Staubli VAL3: HMI_TRAJ.pjx

--- HMI_TRAJ.pjx ---
Parameters version=s8.21Cs9_BS4703 stackSize=5000 millimeterUnit=true
Program file=bind.pgx
Program file=copy.pgx
Program file=deleteItem.pgx
Program file=getTrajID.pgx
Program file=main.pgx
Program file=new.pgx
Program file=onStart.pgx
Program file=refreshlist.pgx
Program file=simulateTRAJ.pgx
Program file=start.pgx
Program file=stop.pgx
Data file=HMI_TRAJ.dtx
Library alias=trajectory path=Disk://source/projectSource/trajectory/trajectory.pjx
Library alias=util path=Disk://HMI_cs9/HMI_util/HMI_util.pjx
Library alias=saveData path=Disk://source/saveData/saveData.pjx
Library alias=HMI_point path=Disk://HMI_cs9/HMI_pointEdit/HMI_pointEdit.pjx
Library alias=simulate path=Disk://HMI_cs9/simulate/simulate.pjx
Library alias=rs path=Disk://source/projectSource/robotStatus/robotStatus.pjx
Type name=trajItem path=Disk://source/template/trajItem/trajItem.pjx

--- HMI_TRAJ.dtx ---
mdesc mNomSpeed
string sUsingLib
string sList
bool bBack
bool bBool[12]
string sPageIndex
string sPageNum
num nPageIndex
num nPageNum
string sNewName
string sFrameList
string sToolList
bool bConfirm
bool bCancel
num nMoveID
string sSelFrame
string sSelTool
string sSelTraj
bool bRefresh
bool bToSave
public trajItem tEditItem
  [0]
    num nFrameIndex
    num nToolIndex
    string sID
    num nMoveID
    pointItem pPointItem
      [0]
        pointRx pPointRx[2]
        jointRx jJointRx
        paraItem pParaItem
          [0]
            mdesc mMdesc
            num nMoveType
            num nActionIndex
            num nPercentage
            ifItem iIfItem
              [0]
                num nSigType[3]
                num nSigIndex[3]
                num nValue[3]
                bool bANDOR[2]
            num nDelay
            num nSigValue
            bool bSafePoint
        string sID
        bool bMarked
        pointRx pInter
string sTrajList
string sTrajList1
string sSessionList
num nIDIsExit

--- main.pgx ---
public program main()
  local bool l_bExit
  local bool l_bResult
  local num l_nSize
  local bool l_bRefresh
begin
  do
    if util:sPage!="traj"
      util:sPage="traj"
      call onStart()
      call bind()
      call util:loadingPage()
      userPage(util:sPage)
      delay(0.5)
    endIf

    if bBool[0]
      bBool[0]=false
      //新建
      call new()
      bRefresh=true
    elseIf bBool[1]
      bBool[1]=false
      //copy
      call copy()
      bRefresh=true
    elseIf bBool[2]
      bBool[2]=false
      //delete
      call deleteItem()
      bRefresh=true
    elseIf bBool[5]
      bBool[5]=false
      call simulateTRAJ(sSelTraj)
      bRefresh=true
    elseIf bBool[6]
      bBool[6]=false
      //编辑
      call trajectory:onSave(bToSave)

      if sSelTraj!=""
        call HMI_point:main(sSelTraj)
      else
        userPageAlert("未选中有效TRAJ")
      endIf
      bRefresh=true

    elseIf bBool[7]
      bBool[7]=false
      //保存
      call trajectory:onSave(bToSave)
      bRefresh=true
    elseIf bBool[8]
      bBool[8]=false
      //head page
      nPageIndex=0
      l_bRefresh=true
    elseIf bBool[9]
      bBool[9]=false
      //page up
      if nPageIndex>0
        nPageIndex=nPageIndex-1
        l_bRefresh=true
      endIf
    elseIf bBool[10]
      bBool[10]=false
      //page down
      if nPageIndex<nPageNum-1
        nPageIndex=nPageIndex+1
        l_bRefresh=true
      endIf
    elseIf bBool[11]
      bBool[11]=false
      //end page
      nPageIndex=nPageNum-1
      l_bRefresh=true
    elseIf bBack
      bBack=false

      call trajectory:onSave(bToSave)

      l_bExit=true
    endIf

    if l_bRefresh or bRefresh
      l_bRefresh=false
      bRefresh=false
      //刷新列表
      call refreshlist()
    endIf
    //jogmode
    call util:jogMode(saveData:nUsingTool,0)

    delay(0)
  until l_bExit==true
end

--- start.pgx ---
program start()
begin
end

--- bind.pgx ---
program bind()
  local num l_i
  local string l_sbtn
begin
  //lbllib
  userPageBind("traj","lbllib","innerHTML",sUsingLib,1,"r")
  //lst
  //  if size(sList)<50
  //    userPageBind("traj","lst1","options",sList,size(sList),"r")
  //    else
  //      popUpMsg("traj数量过大")
  //    endIf
  userPageBind("traj","lst1","value",sSelTraj,1,"rw")
  //button
  userPageBindClick("traj","btnback",bBack,true)
  for l_i = 0 to 11
    l_sbtn="btn"+toString("",l_i)
    userPageBindClick("traj",l_sbtn,bBool[l_i],true)
  endFor

  //page
  userPageBind("traj","lblpageindex","innerHTML",sPageIndex,1,"r")

  userPageBind("traj","lblpagenum","innerHTML",sPageNum,1,"r")


end

--- copy.pgx ---
program copy()
  local string l_sMsg
  local string l_sInputName
  local bool l_bResult
  local bool l_bResult1
  local num l_nID
  local num l_i
  local bool l_bFound
  local num l_nSize
  local string l_sHeader
begin
  l_sMsg="复制"+sSelTraj+"到："
  l_bResult=userPagePrompt(l_sMsg,l_sInputName)
  if l_bResult
    call trajectory:isDefine(l_sInputName,l_bResult1)
    if !l_bResult1
      call trajectory:getSize(l_nSize)
      call getTrajID()
      l_nID=0
      do
        l_i=0
        do
          if l_nID==nIDIsExit[l_i]
            l_bFound=true
            l_nID=l_nID+1
          else
            l_bFound=false
          endIf
          l_i=l_i+1
        until l_bFound==false or l_i>=size(nIDIsExit)

      until l_bFound==false

      if l_nSize<10
        l_sHeader="0"+toString("",l_nID)+" "+l_sInputName
      else
        l_sHeader=toString("",l_nID)+" "+l_sInputName
      endIf

      call trajectory:copy(sSelTraj,l_sHeader,bToSave)
      call trajectory:onSave(bToSave)
    else
      userPageAlert("输入的名称重复！")
    endIf
  endIf
end

--- deleteItem.pgx ---
public program deleteItem()
  local string l_sMsg
  local bool l_bResult
begin
  if sSelTraj!=""
    l_sMsg="是否删除："+sSelTraj+"?"
    l_bResult=userPageConfirm(l_sMsg)
    if l_bResult
      call trajectory:deleteTraj(sSelTraj,bToSave)
      //call trajectory:getTrajList(sList)
    endIf
  else
    userPageAlert("未选中任意项目！")
  endIf
end

--- getTrajID.pgx ---
program getTrajID()
  local num l_nSession
  local num i
  local string l_sEmpty
  local bool l_bOk
begin
  // init
  //  x_bFounded=false
  //  x_sSessionName=""
  //  //
  // get the list
  //
  //  l_sEmpty=""
  call trajectory:getTrajList(sSessionList)
  //
  // search the program from a number:
  //
  // "number+space+name"
  //
  // 01 MyPart
  // 10 YourPart
  //
  resize(nIDIsExit,1,size(sSessionList))
  for i=0 to size(sSessionList)-1
    if sSessionList[i]!=""
      // convert the string "00 name" into a num
      toNum(sSessionList[i],l_nSession,l_bOk)
      if l_bOk
        nIDIsExit[i]=l_nSession
        endIf
    endIf
  endFor
end

--- new.pgx ---
public program new()
  local string l_sPage
  local bool l_bExit
  local num l_i
  local num l_nToolIndex
  local num l_nFrameIndex
  local bool l_bResult
  local bool l_bResult1
  local num l_nSize
  local string l_sHeader
  local num l_nID
  local bool l_bFound
begin
  // l_sPage=""
  do
    if util:sPage!="new"
      util:sPage="new"
      resize(sFrameList,1,size(saveData:fFrameItem))
      resize(sToolList,1,size(saveData:tToolItem))
      for l_i = 0 to size(sFrameList)-1
        sFrameList[l_i]=toString("",l_i)+","+saveData:fFrameItem[l_i].sName
      endFor
      for l_i = 0 to size(sToolList)-1
        sToolList[l_i]=toString("",l_i)+","+saveData:tToolItem[l_i].sName
      endFor
      sNewName=""
      nMoveID=0
      bCancel=false
      bConfirm=false
      sSelFrame=""
      sSelTool=""
      userPageBind("new","txt1","value",sNewName,1,"rw")
      userPageBind("new","nmb1","value",nMoveID,1,"rw")
      userPageBind("new","cbx1","options",sFrameList,size(sFrameList),"r")
      userPageBind("new","cbx2","options",sToolList,size(sToolList),"r")
      userPageBind("new","cbx1","value",sSelFrame,1,"rw")
      userPageBind("new","cbx2","value",sSelTool,1,"rw")
      userPageBindClick("new","btn1",bConfirm,true)
      userPageBindClick("new","btn2",bCancel,true)
      userPage(util:sPage)
      delay(0.5)

    endIf
    //
    toNum(sSelFrame,l_nFrameIndex,l_bResult)
    toNum(sSelTool,l_nToolIndex,l_bResult1)
    //button
    if bConfirm
      bConfirm=false
      if l_bResult and l_bResult1
        call trajectory:getSize(l_nSize)
        call getTrajID()
        l_nID=0
        do
          l_i=0
          do
            if l_nID==nIDIsExit[l_i]
              l_bFound=true
               l_nID=l_nID+1
            else
              l_bFound=false
            endIf
            l_i=l_i+1
          until l_bFound==false or l_i>=size(nIDIsExit)

          until l_bFound==false

        if l_nSize<10
          l_sHeader="0"+toString("",l_nID)+" "+sNewName
        else
          l_sHeader=toString("",l_nID)+" "+sNewName
        endIf
          call trajectory:new(l_sHeader,l_nFrameIndex,l_nToolIndex,nMoveID,bToSave)
          call trajectory:onSave(bToSave)
          sSelTraj=l_sHeader
          l_bExit=true
      else
        popUpMsg("设定的数据非法")
      endIf
    elseIf bCancel
      bCancel=false
      l_bExit=true
    endIf


    delay(0)
  until l_bExit==true

end

--- onStart.pgx ---
program onStart()
  local num l_nResult
  local string l_sKey
  local num l_i
  local num l_nSize
begin

  sUsingLib=toString("",saveData:nLibIndex)
  // l_nResult=trajTemp:libLoad("Disk://data/CustomerLib/lib0/saveTRAJ")
  //  call trajectory:loadTRAJ(0,l_nResult)
  //  if l_nResult!=0
  //    popUpMsg("库加载错误："+toString("",l_nResult))
  //  endIf



  call refreshlist()
  //refresh list
  //  l_sKey=first(trajTemp:tTrajItem)
  //  while l_sKey!=""
  //    sList[size(sList)-1]=l_sKey
  //    insert(sList[size(sList)])
  //    l_sKey=next(trajTemp:tTrajItem[l_sKey])
  //  endWhile

  nPageIndex=0

  if l_nSize>0
    sSelTraj=sList[l_nSize-1]
  else
    sSelTraj=""
  endIf
  //
end

--- refreshlist.pgx ---
program refreshlist()
  local num l_nSize
  local string l_sTrajList
  local num l_i
  local num l_nCount
begin
  call trajectory:getTrajSize(l_nSize)
  call trajectory:getTrajList(sTrajList)
  //page
  if l_nSize<50
    nPageNum=1
  else
    nPageNum=roundUp(l_nSize/49)
  endIf

  //list
  if nPageNum==1
    if l_nSize<1
      for l_i = 0 to size(sList)-1
        sList[l_i]=""
      endFor
    else
      resize(sList,1,l_nSize)
      for l_i = 0 to size(sList)-1
        sList[l_i]=""
      endFor
      for l_i = 0 to l_nSize-1
        sList[l_i]=sTrajList[l_i]
      endFor
    endIf

  else
    if nPageIndex<nPageNum-1
      resize(sList,1,49)
      for l_i = 0 to size(sList)-1
        sList[l_i]=sTrajList[nPageIndex*49+l_i]
      endFor
    else
      for l_i = 0 to size(sList)-1
        sList[l_i]=""
      endFor
      if l_nSize%49==0
        l_nCount=49
      else
        l_nCount=l_nSize%49
      endIf
      resize(sList,1,l_nCount)
      for l_i = 0 to l_nCount-1
        sList[l_i]=sTrajList[l_i+nPageIndex*49]
      endFor
    endIf
  endIf
  userPageBind("traj","lst1","options",sList,size(sList),"r")
  sPageIndex=toString("",nPageIndex+1)
  sPageNum=toString("",nPageNum)
end

--- simulate.pgx ---
program simulate()
begin
end

--- simulateTRAJ.pgx ---
program simulateTRAJ(string x_sKey)
begin
  call simulate:simulateTRAJ(x_sKey)
end

--- stop.pgx ---
program stop()
begin
end
